SUBAPPLICATION Schneidwerk (* Subapplication Type *)
  (* Standard: 61499-2 *)
  (* Version 1.0, 2023-01-29, Franz *)
  IMPORT DefaultPool::SoftKey_Schneidwerk;
  IMPORT isobus::UT::io::Softkey::SoftKeyActivationCode::SK_RELEASED;
  IMPORT DefaultPool::AuxInput_Schneidwerk;
  IMPORT isobus::UT::io::Auxiliary::IN::AuxiliaryState::AuxDisabled;
  IMPORT logiBUS::io::DQ::logiBUS_DO::Output_Q1;
  IMPORT logiBUS::io::DQ::logiBUS_DO::Invalid;
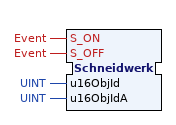
  EVENT_INPUT
    S_ON;
    S_OFF;
  END_EVENT
  VAR_INPUT
    u16ObjId : UINT;
    u16ObjIdA : UINT;
  END_VAR
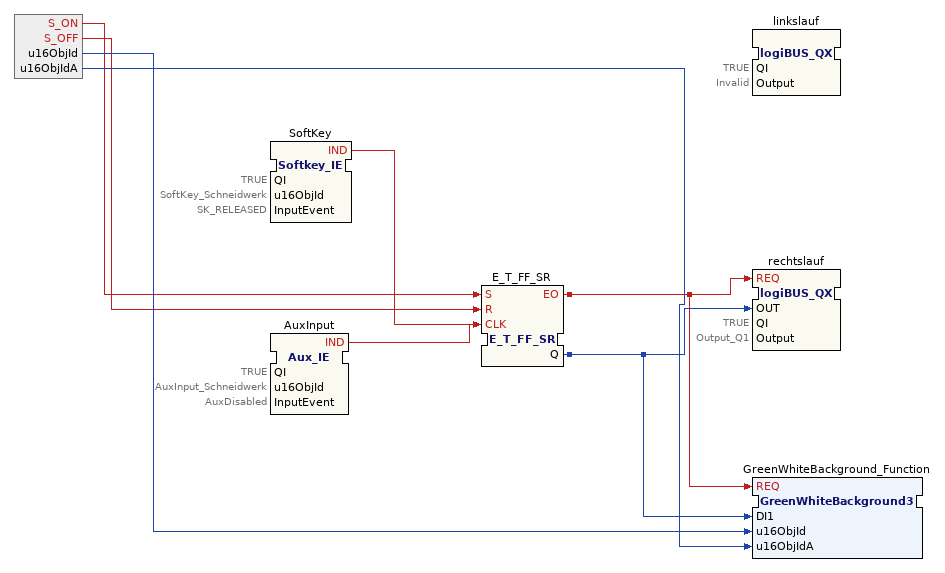
  (* TODO: Schneidwerk linkslauf bei jedem 2. Start. *)
  FBS
    rechtslauf : logiBUS::io::DQ::logiBUS_QX(QI := TRUE, Output := Output_Q1);
    E_T_FF_SR : iec61499::events::E_T_FF_SR;
    linkslauf : logiBUS::io::DQ::logiBUS_QX(QI := TRUE, Output := Invalid);
    SoftKey : isobus::UT::io::Softkey::Softkey_IE(QI := TRUE, u16ObjId := SoftKey_Schneidwerk, InputEvent := SK_RELEASED);
    AuxInput : isobus::UT::io::Auxiliary::IN::Aux_IE(QI := TRUE, u16ObjId := AuxInput_Schneidwerk, InputEvent := AuxDisabled);
  END_FBS
  SUBAPPS
    GreenWhiteBackground_Function : MyLib::sys::GreenWhiteBackground3;
  END_SUBAPPS
  EVENT_CONNECTIONS
    E_T_FF_SR.EO TO rechtslauf.REQ;
    S_ON TO E_T_FF_SR.S;
    S_OFF TO E_T_FF_SR.R;
    E_T_FF_SR.EO TO GreenWhiteBackground_Function.REQ;
    SoftKey.IND TO E_T_FF_SR.CLK;
    AuxInput.IND TO E_T_FF_SR.CLK;
  END_CONNECTIONS
  DATA_CONNECTIONS
    E_T_FF_SR.Q TO rechtslauf.OUT;
    E_T_FF_SR.Q TO GreenWhiteBackground_Function.DI1;
    u16ObjId TO GreenWhiteBackground_Function.u16ObjId;
    u16ObjIdA TO GreenWhiteBackground_Function.u16ObjIdA;
  END_CONNECTIONS
END_SUBAPPLICATION
